Fanuc KAREL source: kx00017.KL

PROGRAM KX00017
%STACKSIZE=65535
%PRIORITY=65535
%NOLOCKGROUP
VAR
I : INTEGER
J : INTEGER
B : BOOLEAN
F : FILE
S : STRING[80]
P : XYZWPR
BEGIN
-- UNRESOLVED_PC line 11 opcodes [03 2E 1B 12 13 04 14] marker_code=0
END KX00017
